TYPE E_ValveState :
(
	Closed := 0,
	Opening := 1,
	Open := 2,
	Closing := 3
);
END_TYPE

(* stored: Version 1.1.0.1, ProductVersion 3.1.4024.12
   DUT E_ValveState: Id {1cc629bf-b40d-4963-adb6-2dda6ec67b55} *)
